(* IEC 61131-3 sources: vscode-twincat-st/src/sample/Complex, 9 files *)

(* ---- Defaults.st ---- *)
VAR_GLOBAL Defaults
	DEFAULT_BOOL: 	BOOL 	:= FALSE;

	DEFAULT_INT: 	INT 	:= 0;

	DEFAULT_REAL: 	REAL	:= 0.0;
END_VAR

(* ---- Periods.st ---- *)
VAR_GLOBAL CONSTANT Periods
	LIFEBIT_TIMEOUT:	TIME := T#10S;

	DEFAULT_DELAY: 		TIME := T#2S;
END_VAR

(* ---- I_Counter.st ---- *)
INTERFACE I_Counter EXTENDS I_CounterBase1, I_CounterBase2
    //
END_INTERFACE

(* ---- I_CounterBase1.st ---- *)
INTERFACE I_CounterBase1

    PROPERTY Value : INT
        GET
            //
        END_GET
        SET
            //
        END_SET
    END_PROPERTY
END_INTERFACE

(* ---- I_CounterBase2.st ---- *)
INTERFACE INTERNAL I_CounterBase2
    //
END_INTERFACE

(* ---- I_Reset.st ---- *)
INTERFACE I_Reset

    METHOD Reset : BOOL
        //
    END_METHOD
END_INTERFACE

(* ---- FB_Counter.st ---- *)
FUNCTION_BLOCK FB_Counter EXTENDS FB_CounterBase IMPLEMENTS I_Counter, I_Reset

    VAR_INPUT
        enable: BOOL := FALSE;

        count:  REFERENCE TO BOOL;

        unused: INT;
    END_VAR

    VAR_OUTPUT
        success: BOOL;
    END_VAR

    VAR
        _value:     INT;
        _unused:    BOOL;
    END_VAR

    PROPERTY Value : INT
        GET
            Value := _value;
        END_GET
        SET
            _value := Value;
        END_SET
    END_PROPERTY

    METHOD Reset : BOOL

        VAR_INST
            _resetCount:    INT;
            _unused:        BOOL;
        END_VAR

        _value      := Defaults.DEFAULT_INT;
        _resetCount := _resetCount MOD 5 + 1;
    END_METHOD

    METHOD PRIVATE UnusedMethod : BOOL
        _value := Defaults.DEFAULT_INT;
    END_METHOD

    METHOD PRIVATE IncreaseByTwo : BOOL
        _value := _value + 1;
    END_METHOD

    IF enable OR FALSE THEN
        THIS^.IncreaseByTwo();
        count := count + 1;
    END_IF;
END_FUNCTION_BLOCK

(* ---- FB_CounterBase.st ---- *)
FUNCTION_BLOCK ABSTRACT FB_CounterBase

    VAR
        _baseInternal: INT;
    END_VAR

    PROPERTY BaseValue : INT
        GET
            BaseValue := _baseInternal;
        END_GET
        SET
            _baseInternal := BaseValue;
        END_SET
    END_PROPERTY

    METHOD ABSTRACT DoSomething : BOOL
        //
    END_METHOD

    METHOD FB_Init

        VAR_INPUT
            bInitRetains : BOOL;
            bInCopyCode  : BOOL;
        END_VAR

        _baseInternal := 0;
    END_METHOD
END_FUNCTION_BLOCK

(* ---- MAIN.st ---- *)
PROGRAM MAIN

    VAR
        _counter:   FB_Counter;
        _enable:    BOOL := TRUE;
        _success:   BOOL;
        _count:     INT;
    END_VAR

    _counter(enable := _enable, count := _count, success => _success);
    _counter.Reset();
    _counter.Value := 99;
END_PROGRAM
